(* IEC 61131-3 sources: sis-interlock-demo/tools/tests/fixtures/lowering/src/POUs/FB_Slots, 4 files *)

(* ---- FB_Slots.decl.st ---- *)
// Назначение: пример для понижения iec-checker (tools/tests/test_assemble.py)
// Автор:      kr0nsch
// Версия:     0.1.0
// Документ:   docs/LAYOUT.md, раздел «Собранный текст build/assembled»; tools/README.md
FUNCTION_BLOCK FB_Slots
VAR_IN_OUT CONSTANT
    stCfg : ST_Cfg;
END_VAR
VAR
    afbDelay : ARRAY[0..GVL_Const.SLOTS_MAX - 1] OF TON;
    aiGrid : ARRAY[0..GRID_LAST, 0..GVL_Const.GRID_MAX] OF INT;
    aaliNested : ARRAY[0..1] OF ARRAY[0..2] OF LINT;
    iSlot : INT;
    xAny : BOOL;
    rSum : REAL;
    wMask : WORD;
    rGain : REAL;
    iState : INT;
END_VAR
VAR CONSTANT
    GRID_LAST : INT := 2;
END_VAR

(* ---- Check.method.decl.st ---- *)
METHOD Check : BOOL
VAR_IN_OUT CONSTANT
    astCfg : ARRAY[0..GVL_Const.SLOTS_MAX - 1] OF ST_Slot;
END_VAR
VAR
    iIdx : INT;
END_VAR

(* ---- Check.method.impl.st ---- *)
Check := TRUE;
FOR iIdx := 0 TO GVL_Const.SLOTS_MAX - 1 DO
    Check := Check AND astCfg[iIdx].rValue >= 0.0;
END_FOR

(* ---- FB_Slots.impl.st ---- *)
// Обращения к элементам массивов, типизированные литералы, AND_THEN и пустые ветви CASE
FOR iSlot := 0 TO GVL_Const.SLOTS_MAX - 1 DO
    afbDelay[iSlot](IN := stCfg.astSlot[iSlot].xEnable, PT := T#1S);
    xAny := xAny OR afbDelay[iSlot].Q;
    rSum := rSum + stCfg.astSlot[iSlot].rValue;
    aiGrid[iSlot, 0] := aiGrid[0, iSlot] + 1;
    aaliNested[0][iSlot] := 0;
END_FOR
wMask := WORD#16#FF;
rGain := REAL#2 * 1E3;  // lint:allow STL008 литерал с экспонентой — пример для понижения
xAny := xAny AND_THEN rSum > 0.0;
CASE iState OF
    0:
    1:
        iState := 2;
ELSE
    ;
END_CASE
Check(astCfg := stCfg.astSlot);
